{attribute 'no_assign'}
FUNCTION_BLOCK FB_LN_WTURBINE_LD0_WMET1 EXTENDS FB_AcsiCommonLogicalNodeClass
VAR_INPUT
	Beh: FB_DO_WTURBINE_LD0_WMET1_Beh := (sClass:='ENS', bLinkResult:=THIS^.AddDataToContainer(ipData:=Beh));
	HorWdDir: FB_DO_WTURBINE_LD0_WMET1_HorWdDir := (sClass:='MV', bLinkResult:=THIS^.AddDataToContainer(ipData:=HorWdDir));
	HorWdSpd: FB_DO_WTURBINE_LD0_WMET1_HorWdSpd := (sClass:='MV', bLinkResult:=THIS^.AddDataToContainer(ipData:=HorWdSpd));
END_VAR
VAR
END_VAR

END_FUNCTION_BLOCK

(* stored: Version 1.1.0.1
   POU FB_LN_WTURBINE_LD0_WMET1: Id {b126cf80-f796-48d4-82e9-0b512aadcfb1}, SpecialFunc None *)
